Fanuc KAREL source: kt00260.KL

-- PROVISIONAL review KL for V940-1; original PC SHA256 c407b03afd28387b2266f7fce3d7af10d3b1ca7a876ea788364ddf27aa26b925
-- Incomplete behavior may be omitted. Consult companion uncertainty JSON. Do not deploy.
PROGRAM KT00260
%NOLOCKGROUP
VAR
  I1 : INTEGER
  OUT : BOOLEAN
-- UNRESOLVED_DECL H2 type=002017
BEGIN
  -- V9_ZERO_TABLE_METADATA_HINT layout=0001; no indexed target words; source/name/runtime held
  -- UNRESOLVED_PC offsets 5-16; opcodes 2E,23
  -- UNRESOLVED_PC offsets 21-35; opcodes 2E,22,9D,33,B4
  -- UNRESOLVED_PC offsets 40-62; opcodes 21,22,9D,33,B3,57,23
  -- UNRESOLVED_PC offsets 67-71; opcodes 7F
END KT00260
